// TIA Portal V20 export
TYPE "WT_IO_Handbedienung _ANA_UDT"
   STRUCT
      iBetriebsart : Int;   // 0=Auto / 1=Hand
      iZustand : Int;   // 0=AUTO / 10=Hand
      rAktuellerWert : Real;
      rHandWert : Real;
      byReserve : Array[0..7] of Byte;
   END_STRUCT;
END_TYPE
